(* IEC 61131-3 sources: vespera/src/POU, 15 files *)

(* ---- F_BuildLinks.st ---- *)
(* Связи "кто на кого подаёт" при заданных положениях клапанов.
   Используется для блокировок (с фактическими положениями) и для определения состава
   маршрутов (с положениями из ROUTE_VALVE). Возвращает число связей. *)
FUNCTION F_BuildLinks : INT
VAR_IN_OUT
    aPos   : ARRAY[1..GVL_Const.N_VALVE] OF INT;
    aLinks : ARRAY[1..GVL_Const.N_LINK] OF ST_Link;
END_VAR
VAR
    n : INT;
END_VAR
VAR CONSTANT
    M : INT := 0;   (* LT_MECH *)
    B : INT := 1;   (* LT_BUNKER *)
    X : INT := 2;   (* LT_INVALID *)
END_VAR

(* ---- приёмное отделение и МУЗ ---- *)
n := n + 1; aLinks[n] := F_Link(GVL_Const.M_GATE1, M, GVL_Const.M_N3, TRUE);
n := n + 1; aLinks[n] := F_Link(GVL_Const.M_N3, B, GVL_Const.B_B4, TRUE);
n := n + 1; aLinks[n] := F_Link(GVL_Const.M_MUZ5_FD, M, GVL_Const.M_MUZ5, TRUE);
n := n + 1; aLinks[n] := F_Link(GVL_Const.M_MUZ5, M, GVL_Const.M_N7, TRUE);
n := n + 1; aLinks[n] := F_Link(GVL_Const.M_MUZ5, M, GVL_Const.M_SH32, FALSE);    (* неиспользуемые отходы 32-31-30 *)
n := n + 1; aLinks[n] := F_Link(GVL_Const.M_MUZ5, M, GVL_Const.M_KC35, FALSE);    (* используемые отходы 35-34 *)
n := n + 1; aLinks[n] := F_Link(GVL_Const.M_MUZ5, M, GVL_Const.M_FAN6, FALSE);
n := n + 1; aLinks[n] := F_Link(GVL_Const.M_FAN6, M, GVL_Const.M_SL6, FALSE);
n := n + 1; aLinks[n] := F_Link(GVL_Const.M_N7, B, GVL_Const.B_B8, TRUE);

(* ---- ТОР-18 ---- *)
n := n + 1; aLinks[n] := F_Link(GVL_Const.M_TOR9_FD, M, GVL_Const.M_TOR9, TRUE);
n := n + 1; aLinks[n] := F_Link(GVL_Const.M_TOR9, M, GVL_Const.M_N11, TRUE);
n := n + 1; aLinks[n] := F_Link(GVL_Const.M_TOR9, M, GVL_Const.M_SH31, FALSE);    (* неиспользуемые 31-30 *)
n := n + 1; aLinks[n] := F_Link(GVL_Const.M_TOR9, M, GVL_Const.M_KC35, FALSE);
n := n + 1; aLinks[n] := F_Link(GVL_Const.M_TOR9, M, GVL_Const.M_FAN10, FALSE);
n := n + 1; aLinks[n] := F_Link(GVL_Const.M_FAN10, M, GVL_Const.M_SL10, FALSE);

(* нория 11 -> 12(1) -> TORBA 13(1) | 12(2) -> БТ | растариватель 15(1) -> нория 16 *)
CASE aPos[GVL_Const.V_V12_1] OF
1:
    n := n + 1; aLinks[n] := F_Link(GVL_Const.M_N11, B, GVL_Const.B_T13_1, TRUE);
2:
    CASE aPos[GVL_Const.V_V12_2] OF
    1:
        n := n + 1; aLinks[n] := F_Link(GVL_Const.M_N11, M, GVL_Const.M_BT14_1, TRUE);
        n := n + 1; aLinks[n] := F_Link(GVL_Const.M_N11, M, GVL_Const.M_BT14_2, TRUE);
    2:
        n := n + 1; aLinks[n] := F_Link(GVL_Const.M_N11, M, GVL_Const.M_N16, TRUE);
    ELSE
        n := n + 1; aLinks[n] := F_Link(GVL_Const.M_N11, X, 0, TRUE);
    END_CASE
ELSE
    n := n + 1; aLinks[n] := F_Link(GVL_Const.M_N11, X, 0, TRUE);
END_CASE

(* ---- блок триерный ---- *)
n := n + 1; aLinks[n] := F_Link(GVL_Const.M_BT14_1, M, GVL_Const.M_N16, TRUE);
n := n + 1; aLinks[n] := F_Link(GVL_Const.M_BT14_2, M, GVL_Const.M_N16, TRUE);
n := n + 1; aLinks[n] := F_Link(GVL_Const.M_BT14_1, M, GVL_Const.M_KC36, FALSE);  (* отходы 36-35-34 *)
n := n + 1; aLinks[n] := F_Link(GVL_Const.M_BT14_2, M, GVL_Const.M_KC36, FALSE);

(* нория 16 -> 12(3) -> бункер 17 (КСП) | нория 20 *)
CASE aPos[GVL_Const.V_V12_3] OF
1:
    n := n + 1; aLinks[n] := F_Link(GVL_Const.M_N16, B, GVL_Const.B_B17, TRUE);
2:
    n := n + 1; aLinks[n] := F_Link(GVL_Const.M_N16, M, GVL_Const.M_N20, TRUE);
ELSE
    n := n + 1; aLinks[n] := F_Link(GVL_Const.M_N16, X, 0, TRUE);
END_CASE

(* ---- КСП-11М ---- *)
n := n + 1; aLinks[n] := F_Link(GVL_Const.M_KSP18_FD, M, GVL_Const.M_KSP18, TRUE);
n := n + 1; aLinks[n] := F_Link(GVL_Const.M_KSP18, M, GVL_Const.M_N20, TRUE);
n := n + 1; aLinks[n] := F_Link(GVL_Const.M_KSP18, M, GVL_Const.M_SH33, FALSE);   (* неиспользуемые 33-31-30 *)
n := n + 1; aLinks[n] := F_Link(GVL_Const.M_KSP18, M, GVL_Const.M_KC35, FALSE);
n := n + 1; aLinks[n] := F_Link(GVL_Const.M_KSP18, M, GVL_Const.M_FAN19, FALSE);
n := n + 1; aLinks[n] := F_Link(GVL_Const.M_FAN19, M, GVL_Const.M_SL19, FALSE);
n := n + 1; aLinks[n] := F_Link(GVL_Const.M_N20, B, GVL_Const.B_B22, TRUE);

(* нория 21 -> 12(4) -> бункер 22 (СП) | Z-нория 26 *)
CASE aPos[GVL_Const.V_V12_4] OF
1:
    n := n + 1; aLinks[n] := F_Link(GVL_Const.M_N21, B, GVL_Const.B_B22, TRUE);
2:
    n := n + 1; aLinks[n] := F_Link(GVL_Const.M_N21, M, GVL_Const.M_ZN26, TRUE);
ELSE
    n := n + 1; aLinks[n] := F_Link(GVL_Const.M_N21, X, 0, TRUE);
END_CASE

(* ---- СП-200 ---- *)
n := n + 1; aLinks[n] := F_Link(GVL_Const.M_SP24_DRV, M, GVL_Const.M_ZN26, TRUE);
n := n + 1; aLinks[n] := F_Link(GVL_Const.M_SP24_DRV, M, GVL_Const.M_KC36, FALSE);
n := n + 1; aLinks[n] := F_Link(GVL_Const.M_SP24_DRV, M, GVL_Const.M_SP24_FAN, FALSE);
n := n + 1; aLinks[n] := F_Link(GVL_Const.M_SP24_FAN, M, GVL_Const.M_FAN25, FALSE);
n := n + 1; aLinks[n] := F_Link(GVL_Const.M_FAN25, M, GVL_Const.M_SL25, FALSE);

(* Z-нория 26 -> выгрузка включена: TORBA 13(2) | выключена: бункер фотосепаратора *)
CASE aPos[GVL_Const.V_V49] OF
1:
    n := n + 1; aLinks[n] := F_Link(GVL_Const.M_ZN26, B, GVL_Const.B_T13_2, TRUE);
2:
    n := n + 1; aLinks[n] := F_Link(GVL_Const.M_ZN26, B, GVL_Const.B_B27, TRUE);
ELSE
    n := n + 1; aLinks[n] := F_Link(GVL_Const.M_ZN26, X, 0, TRUE);
END_CASE

(* ---- фотосепаратор (отходы - напрямую в рамку Биг-Бег) ---- *)
n := n + 1; aLinks[n] := F_Link(GVL_Const.M_FS27, M, GVL_Const.M_ZN29, TRUE);
n := n + 1; aLinks[n] := F_Link(GVL_Const.M_FS27, M, GVL_Const.M_FAN28, FALSE);
n := n + 1; aLinks[n] := F_Link(GVL_Const.M_FAN28, M, GVL_Const.M_SL28, FALSE);
n := n + 1; aLinks[n] := F_Link(GVL_Const.M_ZN29, B, GVL_Const.B_T13_2, TRUE);

(* ---- конвейеры отходов ---- *)
n := n + 1; aLinks[n] := F_Link(GVL_Const.M_SH32, M, GVL_Const.M_SH31, FALSE);
n := n + 1; aLinks[n] := F_Link(GVL_Const.M_SH33, M, GVL_Const.M_SH31, FALSE);
n := n + 1; aLinks[n] := F_Link(GVL_Const.M_SH31, M, GVL_Const.M_SH30, FALSE);
n := n + 1; aLinks[n] := F_Link(GVL_Const.M_KC36, M, GVL_Const.M_KC35, FALSE);
n := n + 1; aLinks[n] := F_Link(GVL_Const.M_KC35, M, GVL_Const.M_KC34, FALSE);

F_BuildLinks := n;
END_FUNCTION

(* ---- F_Link.st ---- *)
FUNCTION F_Link : ST_Link
VAR_INPUT
    iFrom    : INT;
    eTo      : INT;
    iTo      : INT;
    xProduct : BOOL;
END_VAR
F_Link.iFrom := iFrom;
F_Link.eTo := eTo;
F_Link.iTo := iTo;
F_Link.xProduct := xProduct;
END_FUNCTION

(* ---- F_Sec.st ---- *)
(* Секунды (UINT) -> TIME *)
FUNCTION F_Sec : TIME
VAR_INPUT
    uSec : UINT;
END_VAR
F_Sec := UDINT_TO_TIME(UINT_TO_UDINT(uSec) * 1000);
END_FUNCTION

(* ---- F_SyncUint.st ---- *)
(* Уставка в RETAIN <-> регистр панели.
   Если панель изменила регистр (он отличается от последнего выданного значения) -
   принять новое значение с ограничением, затем выдать уставку обратно в регистр. *)
FUNCTION F_SyncUint : BOOL
VAR_INPUT
    uMax : UINT;
END_VAR
VAR_IN_OUT
    uHmi    : UINT;
    uPar    : UINT;
    uShadow : UINT;
END_VAR
IF uHmi <> uShadow THEN
    uPar := MIN(uHmi, uMax);
    F_SyncUint := TRUE;
END_IF
uHmi := uPar;
uShadow := uPar;
END_FUNCTION

(* ---- F_SyncWord.st ---- *)
FUNCTION F_SyncWord : BOOL
VAR_IN_OUT
    wHmi    : WORD;
    wPar    : WORD;
    wShadow : WORD;
END_VAR
IF wHmi <> wShadow THEN
    wPar := wHmi;
    F_SyncWord := TRUE;
END_IF
wHmi := wPar;
wShadow := wPar;
END_FUNCTION

(* ---- FB_Bunker.st ---- *)
(* Бункер с датчиком верхнего уровня. Полный бункер ставит на паузу подающий участок
   маршрута; после освобождения и задержки uTRestart участок запускается снова. *)
FUNCTION_BLOCK FB_Bunker
VAR_INPUT
    xHasSF : BOOL;
    stIn   : ST_BunkerIn;
END_VAR
VAR_IN_OUT
    stHmi : ST_BunkerHmi;
    stPar : ST_BunkerPar;
END_VAR
VAR_OUTPUT
    xFull     : BOOL;
    xAlarm    : BOOL;
    xNewAlarm : BOOL;
END_VAR
VAR
    xDvu      : BOOL;
    wAct      : WORD;
    wAlm      : WORD;
    wSts      : WORD;
    uShDvu    : UINT;
    uShRst    : UINT;
    wShByp    : WORD;
    tonFull   : TON;
    tonClear  : TON;
END_VAR

F_SyncUint(uMax := 600, uHmi := stHmi.uTDvu, uPar := stPar.uTDvu, uShadow := uShDvu);
F_SyncUint(uMax := GVL_Const.T_MAX_S, uHmi := stHmi.uTRestart, uPar := stPar.uTRestart, uShadow := uShRst);
F_SyncWord(wHmi := stHmi.wBypass, wPar := stPar.wBypass, wShadow := wShByp);

xDvu := stIn.xDVU AND (stPar.wBypass AND GVL_Const.BY_DVU) = 0;
tonFull(IN := xDvu, PT := F_Sec(stPar.uTDvu));
tonClear(IN := NOT xDvu, PT := F_Sec(stPar.uTRestart));
IF tonFull.Q THEN
    xFull := TRUE;
ELSIF tonClear.Q THEN
    xFull := FALSE;
END_IF

wAct := 0;
IF xHasSF AND NOT stIn.xSF THEN
    wAct := wAct OR GVL_Const.BA_SF;
END_IF
xNewAlarm := (wAct AND NOT wAlm) <> 0;
IF GVL.xReset THEN
    wAlm := wAct;
ELSE
    wAlm := wAlm OR wAct;
END_IF
xAlarm := wAlm <> 0;

wSts := 0;
IF stIn.xDVU THEN wSts := wSts OR GVL_Const.BS_DVU; END_IF
IF xFull THEN wSts := wSts OR GVL_Const.BS_FULL; END_IF
IF stIn.xDNU THEN wSts := wSts OR GVL_Const.BS_DNU; END_IF
IF (stPar.wBypass AND GVL_Const.BY_DVU) <> 0 THEN wSts := wSts OR GVL_Const.BS_BYPASS; END_IF
IF xAlarm THEN wSts := wSts OR GVL_Const.BS_ALARM; END_IF
stHmi.wSts := wSts;
stHmi.wAlm := wAlm;
END_FUNCTION_BLOCK

(* ---- FB_Mech.st ---- *)
(* Механизм линии: двигатель прямого пуска, привод с ПЧ, заслонка с ПЧ или фотосепаратор.

   Режимы:
   - автомат (MODE_AUTO): работает по требованию маршрута. Пуск после задержки uTOn,
     когда все последующие механизмы уже работают (пуск от последнего к первому).
     Останов после задержки uTOff, когда нет требования и остановились все подающие
     механизмы (останов от первого к последнему);
   - ручной с панели (MODE_MAN): кнопки Пуск/Стоп, пуск разрешён только при работе
     последующих механизмов и неполных бункерах на выходе;
   - местный (MODE_LOCAL): ключ поста в "ручн.", кнопки поста;
   - наладка: ручной режим при GVL.xSetup - без блокировок и датчиков безопасности
     (кроме защит двигателя, аварийного стопа и аварии ПЧ).
   Переход между режимами безударный: команда работы сохраняется. *)
FUNCTION_BLOCK FB_Mech
VAR_INPUT
    stCfg       : ST_MechCfg;
    stIn        : ST_MechIn;
    xDemand     : BOOL;    (* требование активного маршрута *)
    xPredRun    : BOOL;    (* работает подающий механизм - удерживать в работе *)
    xSuccOkAuto : BOOL;    (* все последующие механизмы работают *)
    xSuccOkMan  : BOOL;    (* то же + бункеры на выходе не полны *)
    xPaused     : BOOL;    (* участок на паузе по ДВУ (для индикации) *)
END_VAR
VAR_IN_OUT
    stHmi : ST_MechHmi;
    stPar : ST_MechPar;
END_VAR
VAR_OUTPUT
    stOut     : ST_MechOut;
    xRun      : BOOL;      (* механизм в работе (для блокировок соседних) *)
    xCmd      : BOOL;      (* команда работы *)
    xReady    : BOOL;      (* готов к пуску в маршруте *)
    xAuto     : BOOL;
    xAlarm    : BOOL;
    xNewAlarm : BOOL;      (* появилась новая авария (один цикл) *)
END_VAR
VAR
    eMode      : INT;
    xManualReq : BOOL;
    xSetupNow  : BOOL;
    xStartReq  : BOOL;
    xStopReq   : BOOL;
    xMotorOn   : BOOL;     (* выход на двигатель был включен (предыдущий цикл) *)
    xSeqTrip   : BOOL;
    xSeqLatch  : BOOL;
    wAct       : WORD;
    wAlm       : WORD;
    xToDue     : BOOL;
    xOpened    : BOOL;
    xClosed    : BOOL;
    xGoOpen    : BOOL;
    xGoClose   : BOOL;
    xMoveBlock : BOOL;
    wSts       : WORD;
    uShTOn     : UINT;
    uShTOff    : UINT;
    uShTo      : UINT;
    wShByp     : WORD;
    tonStart   : TON;
    tonStop    : TON;
    tonDksRun  : TON;
    tonDksLost : TON;
    rtDks      : R_TRIG;
    tonDsl1    : TON;
    tonDsl2    : TON;
    tonDp      : TON;
    tonFb      : TON;
    tonMove    : TON;
    tpReset    : TP;
    rtCmd      : R_TRIG;
    ftCmd      : F_TRIG;
    tpOn       : TP;
    tpOff      : TP;
    rtLocStart : R_TRIG;
END_VAR

(* ---- уставки панель <-> RETAIN ---- *)
F_SyncUint(uMax := GVL_Const.T_MAX_S, uHmi := stHmi.uTOn, uPar := stPar.uTOn, uShadow := uShTOn);
F_SyncUint(uMax := GVL_Const.T_MAX_S, uHmi := stHmi.uTOff, uPar := stPar.uTOff, uShadow := uShTOff);
F_SyncUint(uMax := 60000, uHmi := stHmi.uToInterval, uPar := stPar.uToInterval, uShadow := uShTo);
F_SyncWord(wHmi := stHmi.wBypass, wPar := stPar.wBypass, wShadow := wShByp);

(* ---- команды панели ---- *)
xStartReq := (stHmi.wCmd AND GVL_Const.C_START) <> 0;
xStopReq := (stHmi.wCmd AND GVL_Const.C_STOP) <> 0;
IF (stHmi.wCmd AND GVL_Const.C_RESET_TO) <> 0 THEN
    stPar.udSecSinceTO := 0;
END_IF
stHmi.wCmd := stHmi.wCmd AND NOT (GVL_Const.C_START OR GVL_Const.C_STOP OR GVL_Const.C_RESET_TO);

(* механизм, занятый маршрутом, в ручной режим с панели не переводится *)
IF xDemand THEN
    stHmi.wCmd := stHmi.wCmd AND NOT GVL_Const.C_MANUAL;
END_IF
xManualReq := (stHmi.wCmd AND GVL_Const.C_MANUAL) <> 0;

IF stCfg.xHasLocal AND stIn.xLocal THEN
    eMode := GVL_Const.MODE_LOCAL;
ELSIF xManualReq THEN
    eMode := GVL_Const.MODE_MAN;
ELSE
    eMode := GVL_Const.MODE_AUTO;
END_IF
xSetupNow := GVL.xSetup AND eMode = GVL_Const.MODE_MAN;
xAuto := eMode = GVL_Const.MODE_AUTO;

(* ---- аварии ---- *)
wAct := 0;
IF stCfg.xHasQF AND NOT stIn.xQF THEN
    wAct := wAct OR GVL_Const.A_QF;
END_IF

tonDksRun(IN := xMotorOn AND stCfg.eDks <> GVL_Const.DKS_NONE, PT := F_Sec(GVL_Retain.stGlobPar.uTDksGrace));
rtDks(CLK := stIn.xDKS);
IF stCfg.eDks = GVL_Const.DKS_PULSE THEN
    (* таймер перезапускается каждым фронтом импульса *)
    tonDksLost(IN := tonDksRun.Q AND NOT rtDks.Q,
               PT := UDINT_TO_TIME(UINT_TO_UDINT(GVL_Retain.stGlobPar.uTDksPulse) * 100));
ELSE
    tonDksLost(IN := tonDksRun.Q AND NOT stIn.xDKS,
               PT := UDINT_TO_TIME(UINT_TO_UDINT(GVL_Retain.stGlobPar.uTDksPulse) * 100));
END_IF
IF tonDksLost.Q AND (stPar.wBypass AND GVL_Const.BY_DKS) = 0 THEN
    wAct := wAct OR GVL_Const.A_DKS;
END_IF

(* сбег ленты контролируется и на стоящей нории: пуск со сбежавшей лентой запрещён *)
tonDsl1(IN := stCfg.xHasDSL AND NOT stIn.xDSL1, PT := T#1S);
IF tonDsl1.Q AND (stPar.wBypass AND GVL_Const.BY_DSL1) = 0 THEN
    wAct := wAct OR GVL_Const.A_DSL1;
END_IF
tonDsl2(IN := stCfg.xHasDSL AND NOT stIn.xDSL2, PT := T#1S);
IF tonDsl2.Q AND (stPar.wBypass AND GVL_Const.BY_DSL2) = 0 THEN
    wAct := wAct OR GVL_Const.A_DSL2;
END_IF
tonDp(IN := stCfg.xHasDP AND NOT stIn.xDP, PT := T#2S);
IF tonDp.Q AND (stPar.wBypass AND GVL_Const.BY_DP) = 0 THEN
    wAct := wAct OR GVL_Const.A_DP;
END_IF

IF stCfg.xHasEStop AND NOT stIn.xEStop THEN
    wAct := wAct OR GVL_Const.A_ESTOP;
END_IF
(* местный "Стоп" при работе от панели/маршрута: механизм уже отключен аппаратно *)
IF stCfg.xHasLocal AND NOT stIn.xLocStop AND eMode <> GVL_Const.MODE_LOCAL AND (xCmd OR xDemand) THEN
    wAct := wAct OR GVL_Const.A_LOCSTOP;
END_IF

CASE stCfg.eKind OF
GVL_Const.K_FC:
    IF stIn.xFcFault THEN
        wAct := wAct OR GVL_Const.A_FC;
    END_IF
    tonFb(IN := xMotorOn AND NOT stIn.xFcReady, PT := F_Sec(GVL_Retain.stGlobPar.uTFcFb));
    IF tonFb.Q THEN
        wAct := wAct OR GVL_Const.A_FCFB;
    END_IF
GVL_Const.K_GATE:
    IF stIn.xFcFault THEN
        wAct := wAct OR GVL_Const.A_FC;
    END_IF
    tonMove(IN := stOut.qOpen OR stOut.qClose, PT := F_Sec(GVL_Retain.stGlobPar.uTGateMove));
    IF tonMove.Q THEN
        wAct := wAct OR GVL_Const.A_MOVE;
    END_IF
    IF stIn.xFb1 AND stIn.xFb2 THEN
        wAct := wAct OR GVL_Const.A_POS;
    END_IF
GVL_Const.K_FS:
    IF stIn.xErr THEN
        wAct := wAct OR GVL_Const.A_FSERR;
    END_IF
    tonFb(IN := xCmd AND NOT stIn.xFb1, PT := F_Sec(GVL_Retain.stGlobPar.uTFsStart));
    IF tonFb.Q THEN
        wAct := wAct OR GVL_Const.A_FSFB;
    END_IF
END_CASE

IF xSetupNow THEN
    wAct := wAct AND GVL_Const.A_HARD;
END_IF

(* фиксация аварий до сброса *)
xNewAlarm := (wAct AND NOT wAlm) <> 0;
IF GVL.xReset THEN
    wAlm := wAct;
    xSeqLatch := FALSE;
ELSE
    wAlm := wAlm OR wAct;
END_IF
xAlarm := wAlm <> 0;

(* ---- готовность к работе в маршруте ---- *)
xReady := NOT xAlarm AND xAuto AND GVL.xGlobalOk
    AND (NOT stCfg.xHasLocal OR stIn.xLocStop)
    AND (NOT stCfg.xHasEStop OR stIn.xEStop)
    AND (stCfg.eKind <> GVL_Const.K_FS
         OR (stIn.xFb2 AND (stIn.xAux OR (stPar.wBypass AND GVL_Const.BY_AUX) <> 0)));

(* ---- команда работы ---- *)
rtLocStart(CLK := stIn.xLocStart);
CASE eMode OF
GVL_Const.MODE_AUTO:
    tonStart(IN := xDemand AND xSuccOkAuto AND xReady AND NOT xCmd, PT := F_Sec(stPar.uTOn));
    IF tonStart.Q THEN
        xCmd := TRUE;
        xSeqLatch := FALSE;
    END_IF
    tonStop(IN := xCmd AND NOT xDemand AND NOT xPredRun, PT := F_Sec(stPar.uTOff));
    IF tonStop.Q THEN
        xCmd := FALSE;
    END_IF
    xSeqTrip := NOT xSuccOkAuto;

GVL_Const.MODE_MAN:
    tonStart(IN := FALSE);
    tonStop(IN := FALSE);
    IF xStartReq AND NOT xAlarm AND GVL.xGlobalOk AND (xSuccOkMan OR xSetupNow) THEN
        xCmd := TRUE;
        xSeqLatch := FALSE;
    END_IF
    IF xStopReq THEN
        xCmd := FALSE;
    END_IF
    xSeqTrip := NOT xSuccOkMan AND NOT xSetupNow;

GVL_Const.MODE_LOCAL:
    tonStart(IN := FALSE);
    tonStop(IN := FALSE);
    IF rtLocStart.Q AND NOT xAlarm AND stIn.xLocStop THEN
        xCmd := TRUE;
    END_IF
    IF NOT stIn.xLocStop THEN
        xCmd := FALSE;
    END_IF
    xSeqTrip := FALSE;
END_CASE

(* заслонка управляется в местном и ручном режимах кнопками открыть/закрыть, см. ниже *)
IF stCfg.eKind = GVL_Const.K_GATE AND eMode <> GVL_Const.MODE_AUTO THEN
    xCmd := FALSE;
    xSeqTrip := FALSE;
END_IF

IF xCmd AND xSeqTrip THEN
    xSeqLatch := TRUE;
END_IF
(* аварийный стоп, пожар, фазы, отключение цепи управления - останов сразу, без задержек *)
IF xAlarm OR NOT GVL.xGlobalOk OR xSeqTrip THEN
    xCmd := FALSE;
END_IF

(* ---- исполнительная часть ---- *)
stOut.qRun := FALSE;
stOut.qPower := FALSE;
stOut.qOpen := FALSE;
stOut.qClose := FALSE;
stOut.qEnable := FALSE;
tpReset(IN := GVL.xReset, PT := T#1S);
stOut.qReset := tpReset.Q;
rtCmd(CLK := xCmd);
ftCmd(CLK := xCmd);
tpOn(IN := rtCmd.Q AND stCfg.eKind = GVL_Const.K_FS, PT := T#1S);
tpOff(IN := ftCmd.Q AND stCfg.eKind = GVL_Const.K_FS, PT := T#1S);
stOut.qOn := tpOn.Q;
stOut.qOff := tpOff.Q;
xOpened := stIn.xFb1 AND NOT stIn.xFb2;
xClosed := stIn.xFb2 AND NOT stIn.xFb1;

CASE stCfg.eKind OF
GVL_Const.K_DOL:
    stOut.qRun := xCmd;
    xRun := xCmd;
    xMotorOn := xCmd;

GVL_Const.K_FC:
    stOut.qPower := GVL.xSysOn AND (NOT stCfg.xHasQF OR stIn.xQF);
    stOut.qRun := xCmd AND stOut.qPower;
    xRun := stOut.qRun;
    xMotorOn := stOut.qRun;

GVL_Const.K_GATE:
    stOut.qPower := GVL.xSysOn AND (NOT stCfg.xHasQF OR stIn.xQF);
    CASE eMode OF
    GVL_Const.MODE_AUTO:
        xGoOpen := xCmd;
        xGoClose := NOT xCmd;
    GVL_Const.MODE_MAN:
        xGoOpen := (stHmi.wCmd AND GVL_Const.C_OPEN) <> 0 AND (xSuccOkMan OR xSetupNow);
        xGoClose := (stHmi.wCmd AND GVL_Const.C_CLOSE) <> 0;
    ELSE
        xGoOpen := stIn.xLocOpen AND stIn.xLocStop;
        xGoClose := stIn.xLocClose AND stIn.xLocStop;
    END_CASE
    (* при общей аварии заслонка только закрывается - прекращение подачи продукта *)
    xGoOpen := xGoOpen AND GVL.xGlobalOk;
    (* ход прекращается при аварии привода или концевиков до сброса *)
    xMoveBlock := (wAlm AND (GVL_Const.A_QF OR GVL_Const.A_FC OR GVL_Const.A_MOVE OR GVL_Const.A_POS)) <> 0
        OR NOT stOut.qPower;
    stOut.qOpen := xGoOpen AND NOT xGoClose AND NOT xOpened AND NOT xMoveBlock;
    stOut.qClose := xGoClose AND NOT xGoOpen AND NOT xClosed AND NOT xMoveBlock;
    (* проём не закрыт - продукт может поступать на норию *)
    xRun := stOut.qOpen OR xOpened OR (NOT xClosed AND NOT xAlarm);
    xMotorOn := stOut.qOpen OR stOut.qClose;

GVL_Const.K_FS:
    stOut.qEnable := xCmd AND stIn.xFb1;
    xRun := xCmd AND stIn.xFb1;
    xMotorOn := xRun;
END_CASE

(* ---- моточасы ---- *)
IF xMotorOn AND GVL.xPulse1s THEN
    stPar.udSecTotal := stPar.udSecTotal + 1;
    stPar.udSecSinceTO := stPar.udSecSinceTO + 1;
END_IF
stHmi.uHoursTotal := UDINT_TO_UINT(MIN(stPar.udSecTotal / 3600, 65535));
stHmi.uMinutes := UDINT_TO_UINT((stPar.udSecTotal / 60) MOD 60);
stHmi.uHoursSinceTO := UDINT_TO_UINT(MIN(stPar.udSecSinceTO / 3600, 65535));
xToDue := stPar.uToInterval > 0 AND stPar.udSecSinceTO / 3600 >= UINT_TO_UDINT(stPar.uToInterval);

(* ---- состояние для панели ---- *)
wSts := 0;
IF xRun THEN wSts := wSts OR GVL_Const.S_RUN; END_IF
IF xCmd THEN wSts := wSts OR GVL_Const.S_CMD; END_IF
IF xReady THEN wSts := wSts OR GVL_Const.S_READY; END_IF
IF xAlarm THEN wSts := wSts OR GVL_Const.S_ALARM; END_IF
IF eMode = GVL_Const.MODE_LOCAL THEN wSts := wSts OR GVL_Const.S_LOCAL; END_IF
IF eMode = GVL_Const.MODE_MAN THEN wSts := wSts OR GVL_Const.S_MANUAL; END_IF
IF xSetupNow THEN wSts := wSts OR GVL_Const.S_SETUP; END_IF
IF tonStart.IN AND NOT xCmd THEN wSts := wSts OR GVL_Const.S_STARTING; END_IF
IF tonStop.IN THEN wSts := wSts OR GVL_Const.S_STOPPING; END_IF
IF xDemand THEN wSts := wSts OR GVL_Const.S_DEMAND; END_IF
IF xPaused THEN wSts := wSts OR GVL_Const.S_PAUSE; END_IF
IF xToDue THEN wSts := wSts OR GVL_Const.S_TO_DUE; END_IF
IF xOpened THEN wSts := wSts OR GVL_Const.S_OPENED; END_IF
IF xClosed THEN wSts := wSts OR GVL_Const.S_CLOSED; END_IF
IF xSeqLatch THEN wSts := wSts OR GVL_Const.S_SEQ_TRIP; END_IF
IF xSuccOkMan THEN wSts := wSts OR GVL_Const.S_SUCC_OK; END_IF
stHmi.wSts := wSts;
stHmi.wAlm := wAlm;

IF xAlarm THEN
    stHmi.iState := 4;
ELSIF eMode = GVL_Const.MODE_LOCAL THEN
    stHmi.iState := 5;
ELSIF tonStop.IN THEN
    stHmi.iState := 3;
ELSIF xRun THEN
    stHmi.iState := 2;
ELSIF tonStart.IN THEN
    stHmi.iState := 1;
ELSE
    stHmi.iState := 0;
END_IF
END_FUNCTION_BLOCK

(* ---- FB_Valve.st ---- *)
(* Переключатель потока ППМ-2 с электроприводом (поз.12(1)..12(4)) и
   механизм промежуточной выгрузки Z-нории поз.26 (пневмораспределитель 49YA1/49YA2).
   Выход держится до срабатывания датчика положения. Положение задаёт маршрут;
   в ручном режиме - кнопки панели, если подающий механизм стоит. *)
FUNCTION_BLOCK FB_Valve
VAR_INPUT
    xHasSF  : BOOL;
    stIn    : ST_ValveIn;
    iTarget : INT;      (* 0 - нет задания маршрута, 1/2 - положение *)
    xFlow   : BOOL;     (* подающий механизм работает *)
END_VAR
VAR_IN_OUT
    stHmi : ST_ValveHmi;
    stPar : ST_ValvePar;
END_VAR
VAR_OUTPUT
    stOut     : ST_ValveOut;
    iPos      : INT;    (* 0 - не определено, 1, 2 *)
    xReady    : BOOL;
    xAlarm    : BOOL;
    xNewAlarm : BOOL;
END_VAR
VAR
    iGoal    : INT;
    xManual  : BOOL;
    xReq1    : BOOL;
    xReq2    : BOOL;
    xMove1   : BOOL;
    xMove2   : BOOL;
    wAct     : WORD;
    wAlm     : WORD;
    wSts     : WORD;
    uShMove  : UINT;
    tonMove  : TON;
    tofQ1    : TOF;
    tofQ2    : TOF;
END_VAR

F_SyncUint(uMax := 600, uHmi := stHmi.uTMove, uPar := stPar.uTMove, uShadow := uShMove);

IF stIn.xS1 AND NOT stIn.xS2 THEN
    iPos := 1;
ELSIF stIn.xS2 AND NOT stIn.xS1 THEN
    iPos := 2;
ELSE
    iPos := 0;
END_IF

(* ---- аварии ---- *)
wAct := 0;
IF xHasSF AND NOT stIn.xSF THEN
    wAct := wAct OR GVL_Const.VA_SF;
END_IF
tonMove(IN := stOut.q1 OR stOut.q2, PT := F_Sec(stPar.uTMove));
IF tonMove.Q THEN
    wAct := wAct OR GVL_Const.VA_TIMEOUT;
END_IF
IF stIn.xS1 AND stIn.xS2 THEN
    wAct := wAct OR GVL_Const.VA_BOTH;
END_IF
xNewAlarm := (wAct AND NOT wAlm) <> 0;
IF GVL.xReset THEN
    wAlm := wAct;
ELSE
    wAlm := wAlm OR wAct;
END_IF
xAlarm := wAlm <> 0;

(* ---- задание положения ---- *)
IF iTarget <> 0 THEN
    stHmi.wCmd := stHmi.wCmd AND NOT GVL_Const.VC_MANUAL;
END_IF
xManual := (stHmi.wCmd AND GVL_Const.VC_MANUAL) <> 0;
xReq1 := (stHmi.wCmd AND GVL_Const.VC_POS1) <> 0;
xReq2 := (stHmi.wCmd AND GVL_Const.VC_POS2) <> 0;
stHmi.wCmd := stHmi.wCmd AND NOT (GVL_Const.VC_POS1 OR GVL_Const.VC_POS2);

IF iTarget <> 0 THEN
    iGoal := iTarget;
ELSIF xManual THEN
    IF NOT xFlow OR GVL.xSetup THEN
        IF xReq1 THEN
            iGoal := 1;
        ELSIF xReq2 THEN
            iGoal := 2;
        END_IF
    END_IF
ELSE
    iGoal := 0;
END_IF

xMove1 := iGoal = 1 AND iPos <> 1 AND NOT xAlarm AND GVL.xGlobalOk;
xMove2 := iGoal = 2 AND iPos <> 2 AND NOT xAlarm AND GVL.xGlobalOk;
(* пауза 0,5 с при реверсе привода *)
stOut.q1 := xMove1 AND NOT tofQ2.Q;
stOut.q2 := xMove2 AND NOT tofQ1.Q AND NOT stOut.q1;
tofQ1(IN := stOut.q1, PT := T#500MS);
tofQ2(IN := stOut.q2, PT := T#500MS);

xReady := NOT xAlarm AND NOT xManual;

wSts := 0;
IF iPos = 1 THEN wSts := wSts OR GVL_Const.VS_POS1; END_IF
IF iPos = 2 THEN wSts := wSts OR GVL_Const.VS_POS2; END_IF
IF stOut.q1 OR stOut.q2 THEN wSts := wSts OR GVL_Const.VS_MOVING; END_IF
IF xAlarm THEN wSts := wSts OR GVL_Const.VS_ALARM; END_IF
IF xManual THEN wSts := wSts OR GVL_Const.VS_MANUAL; END_IF
IF iTarget <> 0 THEN wSts := wSts OR GVL_Const.VS_ROUTE; END_IF
IF xFlow THEN wSts := wSts OR GVL_Const.VS_FLOW; END_IF
stHmi.wSts := wSts;
stHmi.wAlm := wAlm;
END_FUNCTION_BLOCK

(* ---- PLC_PRG.st ---- *)
(* Главная программа. Вызывается из задачи MAST (циклическая, 20 мс). *)
PROGRAM PLC_PRG

PRG_Inputs();
PRG_System();
PRG_Topology();
PRG_Routes();
PRG_Mechs();
PRG_Outputs();
END_PROGRAM

(* ---- PRG_Inputs.st ---- *)
(* Сгенерировано gen/gen_io.py. Физические входы -> логические сигналы.
   Полярность датчиков - константы CFG_* в GVL_Const. *)
PROGRAM PRG_Inputs

GVL.xSysOnIn := GVL_IO.DI_SYS_ON;
GVL.aEStopIn[1] := GVL_IO.DI_ESTOP_1;
GVL.aEStopIn[2] := GVL_IO.DI_ESTOP_2;
GVL.aEStopIn[3] := GVL_IO.DI_ESTOP_3;
GVL.aEStopIn[4] := GVL_IO.DI_ESTOP_4;
GVL.aEStopIn[5] := GVL_IO.DI_ESTOP_5;
GVL.aEStopIn[6] := GVL_IO.DI_ESTOP_6;
GVL.aEStopIn[7] := GVL_IO.DI_ESTOP_7;
GVL.aEStopIn[8] := GVL_IO.DI_ESTOP_8;
GVL.aEStopIn[9] := GVL_IO.DI_ESTOP_9;
GVL.aEStopIn[10] := GVL_IO.DI_ESTOP_10;
GVL.xFireOkIn := GVL_IO.DI_FIRE_OK;
GVL.xPhaseOkIn := GVL_IO.DI_PHASE_OK;
GVL.aMechIn[GVL_Const.M_N3].xDKS := GVL_IO.DI_N3_DKS;
GVL.aMechIn[GVL_Const.M_N3].xDSL1 := (GVL_IO.DI_N3_DSL1 = GVL_Const.CFG_DSL_OK);
GVL.aMechIn[GVL_Const.M_N3].xDSL2 := (GVL_IO.DI_N3_DSL2 = GVL_Const.CFG_DSL_OK);
GVL.aMechIn[GVL_Const.M_N3].xDP := (GVL_IO.DI_N3_DP = GVL_Const.CFG_DP_OK);
GVL.aMechIn[GVL_Const.M_N3].xLocal := (GVL_IO.DI_N3_SA = GVL_Const.CFG_SA_LOCAL);
GVL.aMechIn[GVL_Const.M_N3].xLocStart := GVL_IO.DI_N3_SB_START;
GVL.aMechIn[GVL_Const.M_N3].xLocStop := GVL_IO.DI_N3_SB_STOP;
GVL.aMechIn[GVL_Const.M_N3].xEStop := GVL_IO.DI_N3_SB_ESTOP;
GVL.aMechIn[GVL_Const.M_N3].xQF := GVL_IO.DI_N3_QF;
GVL.aBunkerIn[GVL_Const.B_B4].xDVU := (GVL_IO.DI_B4_DVU = GVL_Const.CFG_DVU_FULL);
GVL.aBunkerIn[GVL_Const.B_B4].xDNU := (GVL_IO.DI_B4_DNU = GVL_Const.CFG_DNU_ON);
GVL.aMechIn[GVL_Const.M_MUZ5].xQF := GVL_IO.DI_MUZ5_QF;
GVL.aMechIn[GVL_Const.M_MUZ5_FD].xQF := GVL_IO.DI_MUZ5FD_SF;
GVL.aMechIn[GVL_Const.M_MUZ5_FD].xFcFault := (GVL_IO.DI_MUZ5FD_FAULT = GVL_Const.CFG_FC_FAULT);
GVL.aMechIn[GVL_Const.M_MUZ5_FD].xFcReady := GVL_IO.DI_MUZ5FD_READY;
GVL.aMechIn[GVL_Const.M_MUZ5_FD].xEStop := GVL_IO.DI_MUZ5FD_ESTOP;
GVL.aMechIn[GVL_Const.M_FAN6].xQF := GVL_IO.DI_FAN6_QF;
GVL.aMechIn[GVL_Const.M_SL6].xDKS := GVL_IO.DI_SL6_DKS;
GVL.aMechIn[GVL_Const.M_SL6].xQF := GVL_IO.DI_SL6_QF;
GVL.aMechIn[GVL_Const.M_N7].xDKS := GVL_IO.DI_N7_DKS;
GVL.aMechIn[GVL_Const.M_N7].xDSL1 := (GVL_IO.DI_N7_DSL1 = GVL_Const.CFG_DSL_OK);
GVL.aMechIn[GVL_Const.M_N7].xDSL2 := (GVL_IO.DI_N7_DSL2 = GVL_Const.CFG_DSL_OK);
GVL.aMechIn[GVL_Const.M_N7].xDP := (GVL_IO.DI_N7_DP = GVL_Const.CFG_DP_OK);
GVL.aMechIn[GVL_Const.M_N7].xLocal := (GVL_IO.DI_N7_SA = GVL_Const.CFG_SA_LOCAL);
GVL.aMechIn[GVL_Const.M_N7].xLocStart := GVL_IO.DI_N7_SB_START;
GVL.aMechIn[GVL_Const.M_N7].xLocStop := GVL_IO.DI_N7_SB_STOP;
GVL.aMechIn[GVL_Const.M_N7].xEStop := GVL_IO.DI_N7_SB_ESTOP;
GVL.aMechIn[GVL_Const.M_N7].xQF := GVL_IO.DI_N7_QF;
GVL.aBunkerIn[GVL_Const.B_B8].xDVU := (GVL_IO.DI_B8_DVU = GVL_Const.CFG_DVU_FULL);
GVL.aBunkerIn[GVL_Const.B_B8].xDNU := (GVL_IO.DI_B8_DNU = GVL_Const.CFG_DNU_ON);
GVL.aMechIn[GVL_Const.M_TOR9].xQF := GVL_IO.DI_TOR9_QF;
GVL.aMechIn[GVL_Const.M_TOR9_FD].xQF := GVL_IO.DI_TOR9FD_SF;
GVL.aMechIn[GVL_Const.M_TOR9_FD].xFcFault := (GVL_IO.DI_TOR9FD_FAULT = GVL_Const.CFG_FC_FAULT);
GVL.aMechIn[GVL_Const.M_TOR9_FD].xFcReady := GVL_IO.DI_TOR9FD_READY;
GVL.aMechIn[GVL_Const.M_TOR9_FD].xEStop := GVL_IO.DI_TOR9FD_ESTOP;
GVL.aMechIn[GVL_Const.M_FAN10].xQF := GVL_IO.DI_FAN10_QF;
GVL.aMechIn[GVL_Const.M_SL10].xDKS := GVL_IO.DI_SL10_DKS;
GVL.aMechIn[GVL_Const.M_SL10].xQF := GVL_IO.DI_SL10_QF;
GVL.aMechIn[GVL_Const.M_N11].xDKS := GVL_IO.DI_N11_DKS;
GVL.aMechIn[GVL_Const.M_N11].xDSL1 := (GVL_IO.DI_N11_DSL1 = GVL_Const.CFG_DSL_OK);
GVL.aMechIn[GVL_Const.M_N11].xDSL2 := (GVL_IO.DI_N11_DSL2 = GVL_Const.CFG_DSL_OK);
GVL.aMechIn[GVL_Const.M_N11].xDP := (GVL_IO.DI_N11_DP = GVL_Const.CFG_DP_OK);
GVL.aMechIn[GVL_Const.M_N11].xLocal := (GVL_IO.DI_N11_SA = GVL_Const.CFG_SA_LOCAL);
GVL.aMechIn[GVL_Const.M_N11].xLocStart := GVL_IO.DI_N11_SB_START;
GVL.aMechIn[GVL_Const.M_N11].xLocStop := GVL_IO.DI_N11_SB_STOP;
GVL.aMechIn[GVL_Const.M_N11].xEStop := GVL_IO.DI_N11_SB_ESTOP;
GVL.aMechIn[GVL_Const.M_N11].xQF := GVL_IO.DI_N11_QF;
GVL.aValveIn[GVL_Const.V_V12_1].xSF := GVL_IO.DI_V121_SF;
GVL.aValveIn[GVL_Const.V_V12_1].xS1 := GVL_IO.DI_V121_POS1;
GVL.aValveIn[GVL_Const.V_V12_1].xS2 := GVL_IO.DI_V121_POS2;
GVL.aValveIn[GVL_Const.V_V12_2].xSF := GVL_IO.DI_V122_SF;
GVL.aValveIn[GVL_Const.V_V12_2].xS1 := GVL_IO.DI_V122_POS1;
GVL.aValveIn[GVL_Const.V_V12_2].xS2 := GVL_IO.DI_V122_POS2;
GVL.aValveIn[GVL_Const.V_V12_3].xSF := GVL_IO.DI_V123_SF;
GVL.aValveIn[GVL_Const.V_V12_3].xS1 := GVL_IO.DI_V123_POS1;
GVL.aValveIn[GVL_Const.V_V12_3].xS2 := GVL_IO.DI_V123_POS2;
GVL.aValveIn[GVL_Const.V_V12_4].xSF := GVL_IO.DI_V124_SF;
GVL.aValveIn[GVL_Const.V_V12_4].xS1 := GVL_IO.DI_V124_POS1;
GVL.aValveIn[GVL_Const.V_V12_4].xS2 := GVL_IO.DI_V124_POS2;
GVL.aBunkerIn[GVL_Const.B_T13_1].xSF := GVL_IO.DI_T131_SF;
GVL.aBunkerIn[GVL_Const.B_T13_2].xSF := GVL_IO.DI_T132_SF;
GVL.aBunkerIn[GVL_Const.B_T13_1].xDVU := (GVL_IO.DI_T131_DVU = GVL_Const.CFG_DVU_FULL);
GVL.aBunkerIn[GVL_Const.B_T13_1].xDNU := (GVL_IO.DI_T131_DNU = GVL_Const.CFG_DNU_ON);
GVL.aBunkerIn[GVL_Const.B_T13_2].xDVU := (GVL_IO.DI_T132_DVU = GVL_Const.CFG_DVU_FULL);
GVL.aBunkerIn[GVL_Const.B_T13_2].xDNU := (GVL_IO.DI_T132_DNU = GVL_Const.CFG_DNU_ON);
GVL.aMechIn[GVL_Const.M_BT14_1].xQF := GVL_IO.DI_BT141_SF;
GVL.aMechIn[GVL_Const.M_BT14_1].xFcFault := (GVL_IO.DI_BT141_FAULT = GVL_Const.CFG_FC_FAULT);
GVL.aMechIn[GVL_Const.M_BT14_1].xFcReady := GVL_IO.DI_BT141_READY;
GVL.aMechIn[GVL_Const.M_BT14_1].xEStop := GVL_IO.DI_BT14_ESTOP;
GVL.aMechIn[GVL_Const.M_BT14_2].xEStop := GVL_IO.DI_BT14_ESTOP;
GVL.aMechIn[GVL_Const.M_BT14_2].xQF := GVL_IO.DI_BT142_SF;
GVL.aMechIn[GVL_Const.M_BT14_2].xFcFault := (GVL_IO.DI_BT142_FAULT = GVL_Const.CFG_FC_FAULT);
GVL.aMechIn[GVL_Const.M_BT14_2].xFcReady := GVL_IO.DI_BT142_READY;
GVL.aMechIn[GVL_Const.M_N16].xDKS := GVL_IO.DI_N16_DKS;
GVL.aMechIn[GVL_Const.M_N16].xDSL1 := (GVL_IO.DI_N16_DSL1 = GVL_Const.CFG_DSL_OK);
GVL.aMechIn[GVL_Const.M_N16].xDSL2 := (GVL_IO.DI_N16_DSL2 = GVL_Const.CFG_DSL_OK);
GVL.aMechIn[GVL_Const.M_N16].xDP := (GVL_IO.DI_N16_DP = GVL_Const.CFG_DP_OK);
GVL.aMechIn[GVL_Const.M_N16].xLocal := (GVL_IO.DI_N16_SA = GVL_Const.CFG_SA_LOCAL);
GVL.aMechIn[GVL_Const.M_N16].xLocStart := GVL_IO.DI_N16_SB_START;
GVL.aMechIn[GVL_Const.M_N16].xLocStop := GVL_IO.DI_N16_SB_STOP;
GVL.aMechIn[GVL_Const.M_N16].xEStop := GVL_IO.DI_N16_SB_ESTOP;
GVL.aMechIn[GVL_Const.M_N16].xQF := GVL_IO.DI_N16_QF;
GVL.aBunkerIn[GVL_Const.B_B17].xDVU := (GVL_IO.DI_B17_DVU = GVL_Const.CFG_DVU_FULL);
GVL.aBunkerIn[GVL_Const.B_B17].xDNU := (GVL_IO.DI_B17_DNU = GVL_Const.CFG_DNU_ON);
GVL.aMechIn[GVL_Const.M_KSP18].xQF := GVL_IO.DI_KSP18_QF;
GVL.aMechIn[GVL_Const.M_KSP18_FD].xQF := GVL_IO.DI_KSP18FD_SF;
GVL.aMechIn[GVL_Const.M_KSP18_FD].xFcFault := (GVL_IO.DI_KSP18FD_FAULT = GVL_Const.CFG_FC_FAULT);
GVL.aMechIn[GVL_Const.M_KSP18_FD].xFcReady := GVL_IO.DI_KSP18FD_READY;
GVL.aMechIn[GVL_Const.M_KSP18_FD].xEStop := GVL_IO.DI_KSP18FD_ESTOP;
GVL.aMechIn[GVL_Const.M_FAN19].xQF := GVL_IO.DI_FAN19_QF;
GVL.aMechIn[GVL_Const.M_SL19].xDKS := GVL_IO.DI_SL19_DKS;
GVL.aMechIn[GVL_Const.M_SL19].xQF := GVL_IO.DI_SL19_QF;
GVL.aMechIn[GVL_Const.M_N20].xDKS := GVL_IO.DI_N20_DKS;
GVL.aMechIn[GVL_Const.M_N20].xDSL1 := (GVL_IO.DI_N20_DSL1 = GVL_Const.CFG_DSL_OK);
GVL.aMechIn[GVL_Const.M_N20].xDSL2 := (GVL_IO.DI_N20_DSL2 = GVL_Const.CFG_DSL_OK);
GVL.aMechIn[GVL_Const.M_N20].xDP := (GVL_IO.DI_N20_DP = GVL_Const.CFG_DP_OK);
GVL.aMechIn[GVL_Const.M_N20].xLocal := (GVL_IO.DI_N20_SA = GVL_Const.CFG_SA_LOCAL);
GVL.aMechIn[GVL_Const.M_N20].xLocStart := GVL_IO.DI_N20_SB_START;
GVL.aMechIn[GVL_Const.M_N20].xLocStop := GVL_IO.DI_N20_SB_STOP;
GVL.aMechIn[GVL_Const.M_N20].xEStop := GVL_IO.DI_N20_SB_ESTOP;
GVL.aMechIn[GVL_Const.M_N20].xQF := GVL_IO.DI_N20_QF;
GVL.aMechIn[GVL_Const.M_N21].xDKS := GVL_IO.DI_N21_DKS;
GVL.aMechIn[GVL_Const.M_N21].xDSL1 := (GVL_IO.DI_N21_DSL1 = GVL_Const.CFG_DSL_OK);
GVL.aMechIn[GVL_Const.M_N21].xDSL2 := (GVL_IO.DI_N21_DSL2 = GVL_Const.CFG_DSL_OK);
GVL.aMechIn[GVL_Const.M_N21].xDP := (GVL_IO.DI_N21_DP = GVL_Const.CFG_DP_OK);
GVL.aMechIn[GVL_Const.M_N21].xLocal := (GVL_IO.DI_N21_SA = GVL_Const.CFG_SA_LOCAL);
GVL.aMechIn[GVL_Const.M_N21].xLocStart := GVL_IO.DI_N21_SB_START;
GVL.aMechIn[GVL_Const.M_N21].xLocStop := GVL_IO.DI_N21_SB_STOP;
GVL.aMechIn[GVL_Const.M_N21].xEStop := GVL_IO.DI_N21_SB_ESTOP;
GVL.aMechIn[GVL_Const.M_N21].xQF := GVL_IO.DI_N21_QF;
GVL.aBunkerIn[GVL_Const.B_B22].xDVU := (GVL_IO.DI_B22_DVU = GVL_Const.CFG_DVU_FULL);
GVL.aBunkerIn[GVL_Const.B_B22].xDNU := (GVL_IO.DI_B22_DNU = GVL_Const.CFG_DNU_ON);
GVL.aMechIn[GVL_Const.M_SP24_FAN].xQF := GVL_IO.DI_SP24FAN_QF;
GVL.aMechIn[GVL_Const.M_SP24_DRV].xQF := GVL_IO.DI_SP24DRV_SF;
GVL.aMechIn[GVL_Const.M_SP24_DRV].xFcFault := (GVL_IO.DI_SP24DRV_FAULT = GVL_Const.CFG_FC_FAULT);
GVL.aMechIn[GVL_Const.M_SP24_DRV].xFcReady := GVL_IO.DI_SP24DRV_READY;
GVL.aMechIn[GVL_Const.M_SP24_DRV].xEStop := GVL_IO.DI_SP24DRV_ESTOP;
GVL.aMechIn[GVL_Const.M_FAN25].xQF := GVL_IO.DI_FAN25_QF;
GVL.aMechIn[GVL_Const.M_SL25].xDKS := GVL_IO.DI_SL25_DKS;
GVL.aMechIn[GVL_Const.M_SL25].xQF := GVL_IO.DI_SL25_QF;
GVL.aMechIn[GVL_Const.M_FAN28].xQF := GVL_IO.DI_FAN28_QF;
GVL.aMechIn[GVL_Const.M_SL28].xDKS := GVL_IO.DI_SL28_DKS;
GVL.aMechIn[GVL_Const.M_SL28].xQF := GVL_IO.DI_SL28_QF;
GVL.aMechIn[GVL_Const.M_SH31].xDKS := GVL_IO.DI_SH31_DKS;
GVL.aMechIn[GVL_Const.M_SH31].xDP := (GVL_IO.DI_SH31_DP = GVL_Const.CFG_DP_SCREW_OK);
GVL.aMechIn[GVL_Const.M_SH31].xLocal := (GVL_IO.DI_SH31_SA = GVL_Const.CFG_SA_LOCAL);
GVL.aMechIn[GVL_Const.M_SH31].xLocStart := GVL_IO.DI_SH31_SB_START;
GVL.aMechIn[GVL_Const.M_SH31].xLocStop := GVL_IO.DI_SH31_SB_STOP;
GVL.aMechIn[GVL_Const.M_SH31].xEStop := GVL_IO.DI_SH31_SB_END;
GVL.aMechIn[GVL_Const.M_SH31].xQF := GVL_IO.DI_SH31_QF;
GVL.aMechIn[GVL_Const.M_SH32].xDKS := GVL_IO.DI_SH32_DKS;
GVL.aMechIn[GVL_Const.M_SH32].xDP := (GVL_IO.DI_SH32_DP = GVL_Const.CFG_DP_SCREW_OK);
GVL.aMechIn[GVL_Const.M_SH32].xLocal := (GVL_IO.DI_SH32_SA = GVL_Const.CFG_SA_LOCAL);
GVL.aMechIn[GVL_Const.M_SH32].xLocStart := GVL_IO.DI_SH32_SB_START;
GVL.aMechIn[GVL_Const.M_SH32].xLocStop := GVL_IO.DI_SH32_SB_STOP;
GVL.aMechIn[GVL_Const.M_SH32].xEStop := GVL_IO.DI_SH32_SB_END;
GVL.aMechIn[GVL_Const.M_SH32].xQF := GVL_IO.DI_SH32_QF;
GVL.aMechIn[GVL_Const.M_SH33].xDKS := GVL_IO.DI_SH33_DKS;
GVL.aMechIn[GVL_Const.M_SH33].xDP := (GVL_IO.DI_SH33_DP = GVL_Const.CFG_DP_SCREW_OK);
GVL.aMechIn[GVL_Const.M_SH33].xLocal := (GVL_IO.DI_SH33_SA = GVL_Const.CFG_SA_LOCAL);
GVL.aMechIn[GVL_Const.M_SH33].xLocStart := GVL_IO.DI_SH33_SB_START;
GVL.aMechIn[GVL_Const.M_SH33].xLocStop := GVL_IO.DI_SH33_SB_STOP;
GVL.aMechIn[GVL_Const.M_SH33].xEStop := GVL_IO.DI_SH33_SB_END;
GVL.aMechIn[GVL_Const.M_SH33].xQF := GVL_IO.DI_SH33_QF;
GVL.aMechIn[GVL_Const.M_KC34].xDKS := GVL_IO.DI_KC34_DKS;
GVL.aMechIn[GVL_Const.M_KC34].xDP := (GVL_IO.DI_KC34_DP = GVL_Const.CFG_DP_CHAIN_OK);
GVL.aMechIn[GVL_Const.M_KC34].xLocal := (GVL_IO.DI_KC34_SA = GVL_Const.CFG_SA_LOCAL);
GVL.aMechIn[GVL_Const.M_KC34].xLocStart := GVL_IO.DI_KC34_SB_START;
GVL.aMechIn[GVL_Const.M_KC34].xLocStop := GVL_IO.DI_KC34_SB_STOP;
GVL.aMechIn[GVL_Const.M_KC34].xEStop := GVL_IO.DI_KC34_SB_END;
GVL.aMechIn[GVL_Const.M_KC34].xQF := GVL_IO.DI_KC34_QF;
GVL.aMechIn[GVL_Const.M_KC35].xDKS := GVL_IO.DI_KC35_DKS;
GVL.aMechIn[GVL_Const.M_KC35].xDP := (GVL_IO.DI_KC35_DP = GVL_Const.CFG_DP_CHAIN_OK);
GVL.aMechIn[GVL_Const.M_KC35].xLocal := (GVL_IO.DI_KC35_SA = GVL_Const.CFG_SA_LOCAL);
GVL.aMechIn[GVL_Const.M_KC35].xLocStart := GVL_IO.DI_KC35_SB_START;
GVL.aMechIn[GVL_Const.M_KC35].xLocStop := GVL_IO.DI_KC35_SB_STOP;
GVL.aMechIn[GVL_Const.M_KC35].xEStop := GVL_IO.DI_KC35_SB_END;
GVL.aMechIn[GVL_Const.M_KC35].xQF := GVL_IO.DI_KC35_QF;
GVL.aMechIn[GVL_Const.M_KC36].xDKS := GVL_IO.DI_KC36_DKS;
GVL.aMechIn[GVL_Const.M_KC36].xDP := (GVL_IO.DI_KC36_DP = GVL_Const.CFG_DP_CHAIN_OK);
GVL.aMechIn[GVL_Const.M_KC36].xLocal := (GVL_IO.DI_KC36_SA = GVL_Const.CFG_SA_LOCAL);
GVL.aMechIn[GVL_Const.M_KC36].xLocStart := GVL_IO.DI_KC36_SB_START;
GVL.aMechIn[GVL_Const.M_KC36].xLocStop := GVL_IO.DI_KC36_SB_STOP;
GVL.aMechIn[GVL_Const.M_KC36].xEStop := GVL_IO.DI_KC36_SB_END;
GVL.aMechIn[GVL_Const.M_KC36].xQF := GVL_IO.DI_KC36_QF;
GVL.aMechIn[GVL_Const.M_SH30].xDKS := GVL_IO.DI_SH30_DKS;
GVL.aMechIn[GVL_Const.M_SH30].xDP := (GVL_IO.DI_SH30_DP = GVL_Const.CFG_DP_SCREW_OK);
GVL.aMechIn[GVL_Const.M_SH30].xLocal := (GVL_IO.DI_SH30_SA = GVL_Const.CFG_SA_LOCAL);
GVL.aMechIn[GVL_Const.M_SH30].xLocStart := GVL_IO.DI_SH30_SB_START;
GVL.aMechIn[GVL_Const.M_SH30].xLocStop := GVL_IO.DI_SH30_SB_STOP;
GVL.aMechIn[GVL_Const.M_SH30].xEStop := GVL_IO.DI_SH30_SB_END;
GVL.aMechIn[GVL_Const.M_SH30].xQF := GVL_IO.DI_SH30_QF;
GVL.aMechIn[GVL_Const.M_ZN26].xDKS := GVL_IO.DI_ZN26_DKS;
GVL.aMechIn[GVL_Const.M_ZN26].xLocal := (GVL_IO.DI_ZN26_SA = GVL_Const.CFG_SA_LOCAL);
GVL.aMechIn[GVL_Const.M_ZN26].xLocStart := GVL_IO.DI_ZN26_SB_START;
GVL.aMechIn[GVL_Const.M_ZN26].xLocStop := GVL_IO.DI_ZN26_SB_STOP;
GVL.aMechIn[GVL_Const.M_ZN26].xEStop := GVL_IO.DI_ZN26_SB_END;
GVL.aMechIn[GVL_Const.M_ZN26].xFcFault := (GVL_IO.DI_ZN26_FAULT = GVL_Const.CFG_FC_FAULT);
GVL.aMechIn[GVL_Const.M_ZN26].xFcReady := GVL_IO.DI_ZN26_READY;
GVL.aMechIn[GVL_Const.M_ZN26].xQF := GVL_IO.DI_ZN26_SF;
GVL.aValveIn[GVL_Const.V_V49].xS1 := GVL_IO.DI_V49_ON;
GVL.aValveIn[GVL_Const.V_V49].xS2 := GVL_IO.DI_V49_OFF;
GVL.aMechIn[GVL_Const.M_ZN29].xDKS := GVL_IO.DI_ZN29_DKS;
GVL.aMechIn[GVL_Const.M_ZN29].xLocal := (GVL_IO.DI_ZN29_SA = GVL_Const.CFG_SA_LOCAL);
GVL.aMechIn[GVL_Const.M_ZN29].xLocStart := GVL_IO.DI_ZN29_SB_START;
GVL.aMechIn[GVL_Const.M_ZN29].xLocStop := GVL_IO.DI_ZN29_SB_STOP;
GVL.aMechIn[GVL_Const.M_ZN29].xEStop := GVL_IO.DI_ZN29_SB_END;
GVL.aMechIn[GVL_Const.M_ZN29].xFcFault := (GVL_IO.DI_ZN29_FAULT = GVL_Const.CFG_FC_FAULT);
GVL.aMechIn[GVL_Const.M_ZN29].xFcReady := GVL_IO.DI_ZN29_READY;
GVL.aMechIn[GVL_Const.M_ZN29].xQF := GVL_IO.DI_ZN29_SF;
GVL.aMechIn[GVL_Const.M_GATE1].xFb1 := GVL_IO.DI_GATE1_OPENED;
GVL.aMechIn[GVL_Const.M_GATE1].xFb2 := GVL_IO.DI_GATE1_CLOSED;
GVL.aMechIn[GVL_Const.M_GATE1].xLocal := (GVL_IO.DI_GATE1_SA = GVL_Const.CFG_SA_LOCAL);
GVL.aMechIn[GVL_Const.M_GATE1].xLocOpen := GVL_IO.DI_GATE1_SB_OPEN;
GVL.aMechIn[GVL_Const.M_GATE1].xLocClose := GVL_IO.DI_GATE1_SB_CLOSE;
GVL.aMechIn[GVL_Const.M_GATE1].xLocStop := GVL_IO.DI_GATE1_SB_STOP;
GVL.aMechIn[GVL_Const.M_GATE1].xFcFault := (GVL_IO.DI_GATE1_FAULT = GVL_Const.CFG_FC_FAULT);
GVL.aMechIn[GVL_Const.M_GATE1].xFcReady := GVL_IO.DI_GATE1_READY;
GVL.aMechIn[GVL_Const.M_GATE1].xQF := GVL_IO.DI_GATE1_SF;
GVL.aBunkerIn[GVL_Const.B_B27].xDVU := (GVL_IO.DI_B27_DVU1 = GVL_Const.CFG_DVU_FULL);
GVL.aBunkerIn[GVL_Const.B_B27].xDNU := (GVL_IO.DI_B27_DVU2 = GVL_Const.CFG_DNU_ON);
GVL.xFsAspPwrIn := GVL_IO.DI_FS27_ASP_SF;
GVL.aMechIn[GVL_Const.M_FS27].xQF := GVL_IO.DI_FS27_SF;
GVL.aMechIn[GVL_Const.M_FS27].xFb1 := GVL_IO.DI_FS27_STATUS;
GVL.aMechIn[GVL_Const.M_FS27].xFb2 := GVL_IO.DI_FS27_REMOTE;
GVL.aMechIn[GVL_Const.M_FS27].xErr := GVL_IO.DI_FS27_ERROR;
GVL.xDryerOkIn := GVL_IO.DI_DRYER_SF;
GVL.xComprOkIn := GVL_IO.DI_COMPR_SF;
GVL.xCompr2OkIn := GVL_IO.DI_COMPR2_SF;
END_PROGRAM

(* ---- PRG_Mechs.st ---- *)
(* Вызов бункеров, клапанов и механизмов *)
PROGRAM PRG_Mechs
VAR
    i       : INT;
    aBunker : ARRAY[1..GVL_Const.N_BUNKER] OF FB_Bunker;
    aValve  : ARRAY[1..GVL_Const.N_VALVE] OF FB_Valve;
    aMech   : ARRAY[1..GVL_Const.N_MECH] OF FB_Mech;
    xAny    : BOOL;
    xNew    : BOOL;
END_VAR

xAny := FALSE;
xNew := FALSE;

FOR i := 1 TO GVL_Const.N_BUNKER DO
    aBunker[i](xHasSF := GVL_Const.BUNKER_HAS_SF[i],
               stIn := GVL.aBunkerIn[i],
               stHmi := GVL_HMI.aHmiBunker[i],
               stPar := GVL_Retain.aBunkerPar[i]);
    GVL.aBunkerFull[i] := aBunker[i].xFull;
    GVL.aBunkerAlarm[i] := aBunker[i].xAlarm;
    xAny := xAny OR aBunker[i].xAlarm;
    xNew := xNew OR aBunker[i].xNewAlarm;
END_FOR

FOR i := 1 TO GVL_Const.N_VALVE DO
    aValve[i](xHasSF := GVL_Const.VALVE_HAS_SF[i],
              stIn := GVL.aValveIn[i],
              iTarget := GVL.aValveTarget[i],
              xFlow := GVL.aRun[GVL_Const.VALVE_FEEDER[i]],
              stHmi := GVL_HMI.aHmiValve[i],
              stPar := GVL_Retain.aValvePar[i]);
    GVL.aValveOut[i] := aValve[i].stOut;
    GVL.aValvePos[i] := aValve[i].iPos;
    GVL.aValveReady[i] := aValve[i].xReady;
    GVL.aValveAlarm[i] := aValve[i].xAlarm;
    xAny := xAny OR aValve[i].xAlarm;
    xNew := xNew OR aValve[i].xNewAlarm;
END_FOR

FOR i := 1 TO GVL_Const.N_MECH DO
    aMech[i](stCfg := GVL_Const.MECH_CFG[i],
             stIn := GVL.aMechIn[i],
             xDemand := GVL.aDemand[i],
             xPredRun := GVL.aPredRun[i],
             xSuccOkAuto := GVL.aSuccAuto[i],
             xSuccOkMan := GVL.aSuccMan[i],
             xPaused := GVL.aBlocked[i],
             stHmi := GVL_HMI.aHmiMech[i],
             stPar := GVL_Retain.aMechPar[i]);
    GVL.aMechOut[i] := aMech[i].stOut;
    GVL.aRun[i] := aMech[i].xRun;
    GVL.aReady[i] := aMech[i].xReady;
    GVL.aAuto[i] := aMech[i].xAuto;
    GVL.aAlarm[i] := aMech[i].xAlarm;
    xAny := xAny OR aMech[i].xAlarm;
    xNew := xNew OR aMech[i].xNewAlarm;
END_FOR

GVL.xAnyAlarm := xAny;
GVL.xAnyNewAlarm := xNew;
END_PROGRAM

(* ---- PRG_Outputs.st ---- *)
(* Сгенерировано gen/gen_io.py. Логические команды -> физические выходы. *)
PROGRAM PRG_Outputs

GVL_IO.DO_SIREN := GVL.qSiren;
GVL_IO.DO_LAMP_ALARM := GVL.qLamp;
GVL_IO.DO_N3_RUN := GVL.aMechOut[GVL_Const.M_N3].qRun;
GVL_IO.DO_MUZ5_RUN := GVL.aMechOut[GVL_Const.M_MUZ5].qRun;
GVL_IO.DO_MUZ5FD_POWER := GVL.aMechOut[GVL_Const.M_MUZ5_FD].qPower;
GVL_IO.DO_MUZ5FD_RESET := GVL.aMechOut[GVL_Const.M_MUZ5_FD].qReset;
GVL_IO.DO_MUZ5FD_RUN := GVL.aMechOut[GVL_Const.M_MUZ5_FD].qRun;
GVL_IO.DO_FAN6_RUN := GVL.aMechOut[GVL_Const.M_FAN6].qRun;
GVL_IO.DO_SL6_RUN := GVL.aMechOut[GVL_Const.M_SL6].qRun;
GVL_IO.DO_N7_RUN := GVL.aMechOut[GVL_Const.M_N7].qRun;
GVL_IO.DO_TOR9_RUN := GVL.aMechOut[GVL_Const.M_TOR9].qRun;
GVL_IO.DO_TOR9FD_POWER := GVL.aMechOut[GVL_Const.M_TOR9_FD].qPower;
GVL_IO.DO_TOR9FD_RESET := GVL.aMechOut[GVL_Const.M_TOR9_FD].qReset;
GVL_IO.DO_TOR9FD_RUN := GVL.aMechOut[GVL_Const.M_TOR9_FD].qRun;
GVL_IO.DO_FAN10_RUN := GVL.aMechOut[GVL_Const.M_FAN10].qRun;
GVL_IO.DO_SL10_RUN := GVL.aMechOut[GVL_Const.M_SL10].qRun;
GVL_IO.DO_N11_RUN := GVL.aMechOut[GVL_Const.M_N11].qRun;
GVL_IO.DO_V121_POS1 := GVL.aValveOut[GVL_Const.V_V12_1].q1;
GVL_IO.DO_V121_POS2 := GVL.aValveOut[GVL_Const.V_V12_1].q2;
GVL_IO.DO_V122_POS1 := GVL.aValveOut[GVL_Const.V_V12_2].q1;
GVL_IO.DO_V122_POS2 := GVL.aValveOut[GVL_Const.V_V12_2].q2;
GVL_IO.DO_V123_POS1 := GVL.aValveOut[GVL_Const.V_V12_3].q1;
GVL_IO.DO_V123_POS2 := GVL.aValveOut[GVL_Const.V_V12_3].q2;
GVL_IO.DO_V124_POS1 := GVL.aValveOut[GVL_Const.V_V12_4].q1;
GVL_IO.DO_V124_POS2 := GVL.aValveOut[GVL_Const.V_V12_4].q2;
GVL_IO.DO_A18_Q9_RES := FALSE;
GVL_IO.DO_BT141_POWER := GVL.aMechOut[GVL_Const.M_BT14_1].qPower;
GVL_IO.DO_BT141_RESET := GVL.aMechOut[GVL_Const.M_BT14_1].qReset;
GVL_IO.DO_BT141_RUN := GVL.aMechOut[GVL_Const.M_BT14_1].qRun;
GVL_IO.DO_BT142_POWER := GVL.aMechOut[GVL_Const.M_BT14_2].qPower;
GVL_IO.DO_BT142_RESET := GVL.aMechOut[GVL_Const.M_BT14_2].qReset;
GVL_IO.DO_BT142_RUN := GVL.aMechOut[GVL_Const.M_BT14_2].qRun;
GVL_IO.DO_N16_RUN := GVL.aMechOut[GVL_Const.M_N16].qRun;
GVL_IO.DO_KSP18_RUN := GVL.aMechOut[GVL_Const.M_KSP18].qRun;
GVL_IO.DO_KSP18FD_POWER := GVL.aMechOut[GVL_Const.M_KSP18_FD].qPower;
GVL_IO.DO_KSP18FD_RESET := GVL.aMechOut[GVL_Const.M_KSP18_FD].qReset;
GVL_IO.DO_KSP18FD_RUN := GVL.aMechOut[GVL_Const.M_KSP18_FD].qRun;
GVL_IO.DO_FAN19_RUN := GVL.aMechOut[GVL_Const.M_FAN19].qRun;
GVL_IO.DO_SL19_RUN := GVL.aMechOut[GVL_Const.M_SL19].qRun;
GVL_IO.DO_N20_RUN := GVL.aMechOut[GVL_Const.M_N20].qRun;
GVL_IO.DO_N21_RUN := GVL.aMechOut[GVL_Const.M_N21].qRun;
GVL_IO.DO_SP24FAN_RUN := GVL.aMechOut[GVL_Const.M_SP24_FAN].qRun;
GVL_IO.DO_SP24DRV_POWER := GVL.aMechOut[GVL_Const.M_SP24_DRV].qPower;
GVL_IO.DO_SP24DRV_RESET := GVL.aMechOut[GVL_Const.M_SP24_DRV].qReset;
GVL_IO.DO_SP24DRV_RUN := GVL.aMechOut[GVL_Const.M_SP24_DRV].qRun;
GVL_IO.DO_FAN25_RUN := GVL.aMechOut[GVL_Const.M_FAN25].qRun;
GVL_IO.DO_SL25_RUN := GVL.aMechOut[GVL_Const.M_SL25].qRun;
GVL_IO.DO_FAN28_RUN := GVL.aMechOut[GVL_Const.M_FAN28].qRun;
GVL_IO.DO_SL28_RUN := GVL.aMechOut[GVL_Const.M_SL28].qRun;
GVL_IO.DO_SH31_RUN := GVL.aMechOut[GVL_Const.M_SH31].qRun;
GVL_IO.DO_SH32_RUN := GVL.aMechOut[GVL_Const.M_SH32].qRun;
GVL_IO.DO_SH33_RUN := GVL.aMechOut[GVL_Const.M_SH33].qRun;
GVL_IO.DO_KC34_RUN := GVL.aMechOut[GVL_Const.M_KC34].qRun;
GVL_IO.DO_KC35_RUN := GVL.aMechOut[GVL_Const.M_KC35].qRun;
GVL_IO.DO_KC36_RUN := GVL.aMechOut[GVL_Const.M_KC36].qRun;
GVL_IO.DO_SH30_RUN := GVL.aMechOut[GVL_Const.M_SH30].qRun;
GVL_IO.DO_ZN26_POWER := GVL.aMechOut[GVL_Const.M_ZN26].qPower;
GVL_IO.DO_ZN26_RUN := GVL.aMechOut[GVL_Const.M_ZN26].qRun;
GVL_IO.DO_ZN26_RESET := GVL.aMechOut[GVL_Const.M_ZN26].qReset;
GVL_IO.DO_V49_ON := GVL.aValveOut[GVL_Const.V_V49].q1;
GVL_IO.DO_V49_OFF := GVL.aValveOut[GVL_Const.V_V49].q2;
GVL_IO.DO_ZN29_POWER := GVL.aMechOut[GVL_Const.M_ZN29].qPower;
GVL_IO.DO_ZN29_RUN := GVL.aMechOut[GVL_Const.M_ZN29].qRun;
GVL_IO.DO_ZN29_RESET := GVL.aMechOut[GVL_Const.M_ZN29].qReset;
GVL_IO.DO_GATE1_POWER := GVL.aMechOut[GVL_Const.M_GATE1].qPower;
GVL_IO.DO_GATE1_OPEN := GVL.aMechOut[GVL_Const.M_GATE1].qOpen;
GVL_IO.DO_GATE1_RESET := GVL.aMechOut[GVL_Const.M_GATE1].qReset;
GVL_IO.DO_GATE1_CLOSE := GVL.aMechOut[GVL_Const.M_GATE1].qClose;
GVL_IO.DO_FS27_ON := GVL.aMechOut[GVL_Const.M_FS27].qOn;
GVL_IO.DO_FS27_OFF := GVL.aMechOut[GVL_Const.M_FS27].qOff;
GVL_IO.DO_FS27_ENABLE := GVL.aMechOut[GVL_Const.M_FS27].qEnable;
GVL_IO.DO_A19_Q23_RES := FALSE;
GVL_IO.DO_A19_Q24_RES := FALSE;
END_PROGRAM

(* ---- PRG_Routes.st ---- *)
(* Маршруты (Приложение 5). Пуск: проверка готовности -> предпусковой сигнал ->
   перевод клапанов -> работа (механизмы запускаются от последнего к первому).
   Стоп: снятие требования (останов от первого к последнему с задержками).
   Авария механизма/клапана/бункера маршрута или общая авария - останов маршрута. *)
PROGRAM PRG_Routes
VAR
    xInit     : BOOL;
    r         : INT;
    p         : INT;
    i         : INT;
    v         : INT;
    b         : INT;
    h         : INT;
    k         : INT;
    nL        : INT;
    aPosT     : ARRAY[1..GVL_Const.N_VALVE] OF INT;
    aL        : ARRAY[1..GVL_Const.N_LINK] OF ST_Link;
    aTonPre   : ARRAY[1..GVL_Const.N_ROUTE] OF TON;
    xToggle   : BOOL;
    xStop     : BOOL;
    xConflict : BOOL;
    xFault    : BOOL;
    xBusy     : BOOL;
    xShared   : BOOL;
    xPaused   : BOOL;
    xAllRun   : BOOL;
    xValvesOk : BOOL;
    iBad      : INT;
    wSts      : WORD;
    aNotReady : ARRAY[1..GVL_Const.N_ROUTE] OF BOOL;
END_VAR

(* ---- состав маршрутов: обход связей от головных механизмов при положениях клапанов маршрута ---- *)
IF NOT xInit THEN
    FOR r := 1 TO GVL_Const.N_ROUTE DO
        FOR v := 1 TO GVL_Const.N_VALVE DO
            aPosT[v] := GVL_Const.ROUTE_VALVE[r, v];
        END_FOR
        nL := F_BuildLinks(aPos := aPosT, aLinks := aL);
        FOR i := 1 TO GVL_Const.N_MECH DO
            GVL.aMember[r, i] := FALSE;
        END_FOR
        FOR b := 1 TO GVL_Const.N_BUNKER DO
            GVL.aMemberB[r, b] := FALSE;
        END_FOR
        GVL.aRouteCfgErr[r] := FALSE;
        FOR h := 1 TO GVL_Const.N_HEAD DO
            IF GVL_Const.ROUTE_HEAD[r, h] > 0 THEN
                GVL.aMember[r, GVL_Const.ROUTE_HEAD[r, h]] := TRUE;
            END_IF
        END_FOR
        FOR p := 1 TO GVL_Const.N_MECH DO
            FOR k := 1 TO nL DO
                IF GVL.aMember[r, aL[k].iFrom] THEN
                    CASE aL[k].eTo OF
                    GVL_Const.LT_MECH:
                        GVL.aMember[r, aL[k].iTo] := TRUE;
                    GVL_Const.LT_BUNKER:
                        GVL.aMemberB[r, aL[k].iTo] := TRUE;
                    ELSE
                        GVL.aRouteCfgErr[r] := TRUE;
                    END_CASE
                END_IF
            END_FOR
        END_FOR
    END_FOR
    xInit := TRUE;
END_IF

FOR r := 1 TO GVL_Const.N_ROUTE DO
    xToggle := (GVL_HMI.aHmiRoute[r].wCmd AND GVL_Const.RC_TOGGLE) <> 0;
    xStop := (GVL_HMI.aHmiRoute[r].wCmd AND GVL_Const.RC_STOP) <> 0 OR GVL.xStopAll;
    GVL_HMI.aHmiRoute[r].wCmd := 0;

    xConflict := FALSE;
    FOR p := 1 TO GVL_Const.N_ROUTE DO
        IF p <> r AND GVL_Const.ROUTE_CONFLICT[r, p] AND GVL.aRouteState[p] <> GVL_Const.RST_IDLE THEN
            xConflict := TRUE;
        END_IF
    END_FOR

    xValvesOk := TRUE;
    FOR v := 1 TO GVL_Const.N_VALVE DO
        IF GVL_Const.ROUTE_VALVE[r, v] <> 0 AND GVL.aValvePos[v] <> GVL_Const.ROUTE_VALVE[r, v] THEN
            xValvesOk := FALSE;
        END_IF
    END_FOR

    (* ---- контроль аварий активного маршрута ---- *)
    IF GVL.aRouteState[r] <> GVL_Const.RST_IDLE AND GVL.aRouteState[r] <> GVL_Const.RST_STOPPING THEN
        xFault := NOT GVL.xGlobalOk;
        FOR i := 1 TO GVL_Const.N_MECH DO
            IF GVL.aMember[r, i] AND (GVL.aAlarm[i] OR NOT GVL.aAuto[i]) THEN
                xFault := TRUE;
            END_IF
        END_FOR
        FOR v := 1 TO GVL_Const.N_VALVE DO
            IF GVL_Const.ROUTE_VALVE[r, v] <> 0 AND GVL.aValveAlarm[v] THEN
                xFault := TRUE;
            END_IF
        END_FOR
        FOR b := 1 TO GVL_Const.N_BUNKER DO
            IF GVL.aMemberB[r, b] AND GVL.aBunkerAlarm[b] THEN
                xFault := TRUE;
            END_IF
        END_FOR
        IF GVL.aRouteState[r] = GVL_Const.RST_RUN AND NOT xValvesOk THEN
            xFault := TRUE;
        END_IF
        IF xFault THEN
            GVL.aRouteFault[r] := TRUE;
            GVL.aRouteState[r] := GVL_Const.RST_STOPPING;
        END_IF
    END_IF

    CASE GVL.aRouteState[r] OF
    GVL_Const.RST_IDLE:
        IF GVL.xReset THEN
            GVL.aRouteFault[r] := FALSE;
            aNotReady[r] := FALSE;
        END_IF
        IF xToggle THEN
            iBad := 0;
            IF NOT GVL.xGlobalOk THEN
                iBad := -1;
            ELSIF xConflict THEN
                iBad := -2;
            ELSIF GVL.aRouteCfgErr[r] THEN
                iBad := -3;
            ELSE
                FOR i := GVL_Const.N_MECH TO 1 BY -1 DO
                    IF GVL.aMember[r, i] AND NOT GVL.aReady[i] THEN
                        iBad := i;
                    END_IF
                END_FOR
                IF iBad = 0 THEN
                    FOR v := GVL_Const.N_VALVE TO 1 BY -1 DO
                        IF GVL_Const.ROUTE_VALVE[r, v] <> 0 AND NOT GVL.aValveReady[v] THEN
                            iBad := 100 + v;
                        END_IF
                    END_FOR
                END_IF
                IF iBad = 0 THEN
                    FOR b := GVL_Const.N_BUNKER TO 1 BY -1 DO
                        IF GVL.aMemberB[r, b] AND GVL.aBunkerAlarm[b] THEN
                            iBad := 200 + b;
                        END_IF
                    END_FOR
                END_IF
            END_IF
            GVL_HMI.aHmiRoute[r].iNotReady := iBad;
            aNotReady[r] := iBad <> 0;
            IF iBad = 0 THEN
                GVL.aRouteFault[r] := FALSE;
                GVL.aRouteState[r] := GVL_Const.RST_PRESTART;
            END_IF
        END_IF

    GVL_Const.RST_PRESTART:
        IF xStop OR xToggle THEN
            GVL.aRouteState[r] := GVL_Const.RST_IDLE;
        ELSIF aTonPre[r].Q THEN
            GVL.aRouteState[r] := GVL_Const.RST_VALVES;
        END_IF

    GVL_Const.RST_VALVES:
        IF xStop OR xToggle THEN
            GVL.aRouteState[r] := GVL_Const.RST_STOPPING;
        ELSIF xValvesOk THEN
            GVL.aRouteState[r] := GVL_Const.RST_RUN;
        END_IF

    GVL_Const.RST_RUN:
        IF xStop OR xToggle THEN
            GVL.aRouteState[r] := GVL_Const.RST_STOPPING;
        END_IF

    GVL_Const.RST_STOPPING:
        (* ждать останова всех механизмов маршрута, кроме занятых другим работающим маршрутом *)
        xBusy := FALSE;
        FOR i := 1 TO GVL_Const.N_MECH DO
            IF GVL.aMember[r, i] AND GVL.aRun[i] THEN
                xShared := FALSE;
                FOR p := 1 TO GVL_Const.N_ROUTE DO
                    IF p <> r AND GVL.aRouteState[p] = GVL_Const.RST_RUN AND GVL.aMember[p, i] THEN
                        xShared := TRUE;
                    END_IF
                END_FOR
                IF NOT xShared THEN
                    xBusy := TRUE;
                END_IF
            END_IF
        END_FOR
        IF NOT xBusy THEN
            GVL.aRouteState[r] := GVL_Const.RST_IDLE;
        END_IF
    END_CASE

    aTonPre[r](IN := GVL.aRouteState[r] = GVL_Const.RST_PRESTART,
               PT := F_Sec(GVL_Retain.stGlobPar.uTPreStart));
END_FOR

(* ---- требования к механизмам и клапанам ---- *)
FOR i := 1 TO GVL_Const.N_MECH DO
    GVL.aDemand[i] := FALSE;
    FOR r := 1 TO GVL_Const.N_ROUTE DO
        IF GVL.aRouteState[r] = GVL_Const.RST_RUN AND GVL.aMember[r, i] THEN
            GVL.aDemand[i] := TRUE;
        END_IF
    END_FOR
    GVL.aDemand[i] := GVL.aDemand[i] AND NOT GVL.aBlocked[i];
END_FOR

GVL.xPreStart := FALSE;
FOR v := 1 TO GVL_Const.N_VALVE DO
    GVL.aValveTarget[v] := 0;
END_FOR
FOR r := 1 TO GVL_Const.N_ROUTE DO
    IF GVL.aRouteState[r] = GVL_Const.RST_PRESTART THEN
        GVL.xPreStart := TRUE;
    END_IF
    IF GVL.aRouteState[r] <> GVL_Const.RST_IDLE THEN
        FOR v := 1 TO GVL_Const.N_VALVE DO
            IF GVL_Const.ROUTE_VALVE[r, v] <> 0 THEN
                GVL.aValveTarget[v] := GVL_Const.ROUTE_VALVE[r, v];
            END_IF
        END_FOR
    END_IF
END_FOR

(* ---- состояние для панели ---- *)
FOR r := 1 TO GVL_Const.N_ROUTE DO
    xConflict := FALSE;
    FOR p := 1 TO GVL_Const.N_ROUTE DO
        IF p <> r AND GVL_Const.ROUTE_CONFLICT[r, p] AND GVL.aRouteState[p] <> GVL_Const.RST_IDLE THEN
            xConflict := TRUE;
        END_IF
    END_FOR
    xPaused := FALSE;
    xAllRun := GVL.aRouteState[r] = GVL_Const.RST_RUN;
    FOR i := 1 TO GVL_Const.N_MECH DO
        IF GVL.aMember[r, i] THEN
            IF GVL.aBlocked[i] THEN
                xPaused := TRUE;
            ELSIF NOT GVL.aRun[i] THEN
                xAllRun := FALSE;
            END_IF
        END_IF
    END_FOR
    wSts := 0;
    IF GVL.aRouteState[r] <> GVL_Const.RST_IDLE THEN wSts := wSts OR GVL_Const.RS_ACTIVE; END_IF
    IF GVL.aRouteState[r] = GVL_Const.RST_PRESTART THEN wSts := wSts OR GVL_Const.RS_PRESTART; END_IF
    IF GVL.aRouteState[r] = GVL_Const.RST_VALVES THEN wSts := wSts OR GVL_Const.RS_VALVES; END_IF
    IF GVL.aRouteState[r] = GVL_Const.RST_RUN THEN wSts := wSts OR GVL_Const.RS_RUN; END_IF
    IF GVL.aRouteState[r] = GVL_Const.RST_STOPPING THEN wSts := wSts OR GVL_Const.RS_STOPPING; END_IF
    IF xPaused AND GVL.aRouteState[r] = GVL_Const.RST_RUN THEN wSts := wSts OR GVL_Const.RS_PAUSED; END_IF
    IF GVL.aRouteFault[r] THEN wSts := wSts OR GVL_Const.RS_FAULT; END_IF
    IF aNotReady[r] THEN wSts := wSts OR GVL_Const.RS_NOTREADY; END_IF
    IF xConflict THEN wSts := wSts OR GVL_Const.RS_CONFLICT; END_IF
    IF xAllRun THEN wSts := wSts OR GVL_Const.RS_ALLRUN; END_IF
    GVL_HMI.aHmiRoute[r].wSts := wSts;
    GVL_HMI.aHmiRoute[r].iState := GVL.aRouteState[r];
END_FOR
END_PROGRAM

(* ---- PRG_System.st ---- *)
(* Общие сигналы: цепь управления, аварийные стопы, пожар, контроль фаз, сброс, наладка,
   сирена и лампа "Авария", секундный импульс, уставки по умолчанию. *)
PROGRAM PRG_System
VAR
    i         : INT;
    wAct      : WORD;
    wAlm      : WORD;
    wWarn     : WORD;
    wSts      : WORD;
    xNewG     : BOOL;
    xSirenLatch : BOOL;
    tonSec    : TON;
    tonBlink  : TON;
    xBlinkReq : BOOL;
    uSh       : ARRAY[1..7] OF UINT;
END_VAR

(* ---- уставки по умолчанию при первом запуске / потере RETAIN ---- *)
IF GVL_Retain.uInitMagic <> GVL_Const.RETAIN_MAGIC THEN
    GVL_Retain.stGlobPar.uTPreStart := 10;
    GVL_Retain.stGlobPar.uTDksGrace := 5;
    GVL_Retain.stGlobPar.uTDksPulse := 30;
    GVL_Retain.stGlobPar.uTFcFb := 5;
    GVL_Retain.stGlobPar.uTFsStart := 60;
    GVL_Retain.stGlobPar.uTGateMove := 90;
    GVL_Retain.stGlobPar.uSirenOn := 1;
    FOR i := 1 TO GVL_Const.N_MECH DO
        GVL_Retain.aMechPar[i].uTOn := GVL_Const.MECH_CFG[i].uDefTOn;
        GVL_Retain.aMechPar[i].uTOff := GVL_Const.MECH_CFG[i].uDefTOff;
        GVL_Retain.aMechPar[i].uToInterval := 0;
        GVL_Retain.aMechPar[i].wBypass := 0;
    END_FOR
    FOR i := 1 TO GVL_Const.N_VALVE DO
        GVL_Retain.aValvePar[i].uTMove := 30;
    END_FOR
    FOR i := 1 TO GVL_Const.N_BUNKER DO
        GVL_Retain.aBunkerPar[i].wBypass := 0;
        GVL_Retain.aBunkerPar[i].uTDvu := 3;
        GVL_Retain.aBunkerPar[i].uTRestart := 30;
    END_FOR
    GVL_Retain.uInitMagic := GVL_Const.RETAIN_MAGIC;
END_IF

F_SyncUint(uMax := 600, uHmi := GVL_HMI.stHmiG.uTPreStart, uPar := GVL_Retain.stGlobPar.uTPreStart, uShadow := uSh[1]);
F_SyncUint(uMax := 600, uHmi := GVL_HMI.stHmiG.uTDksGrace, uPar := GVL_Retain.stGlobPar.uTDksGrace, uShadow := uSh[2]);
F_SyncUint(uMax := 600, uHmi := GVL_HMI.stHmiG.uTDksPulse, uPar := GVL_Retain.stGlobPar.uTDksPulse, uShadow := uSh[3]);
F_SyncUint(uMax := 600, uHmi := GVL_HMI.stHmiG.uTFcFb, uPar := GVL_Retain.stGlobPar.uTFcFb, uShadow := uSh[4]);
F_SyncUint(uMax := 600, uHmi := GVL_HMI.stHmiG.uTFsStart, uPar := GVL_Retain.stGlobPar.uTFsStart, uShadow := uSh[5]);
F_SyncUint(uMax := 600, uHmi := GVL_HMI.stHmiG.uTGateMove, uPar := GVL_Retain.stGlobPar.uTGateMove, uShadow := uSh[6]);
F_SyncUint(uMax := 1, uHmi := GVL_HMI.stHmiG.uSirenOn, uPar := GVL_Retain.stGlobPar.uSirenOn, uShadow := uSh[7]);

(* ---- такты ---- *)
tonSec(IN := NOT tonSec.Q, PT := T#1S);
GVL.xPulse1s := tonSec.Q;
tonBlink(IN := NOT tonBlink.Q, PT := T#500MS);
IF tonBlink.Q THEN
    xBlinkReq := NOT xBlinkReq;
END_IF
GVL.xBlink := xBlinkReq;
IF GVL.xPulse1s THEN
    GVL_HMI.stHmiG.uHeartbeat := GVL_HMI.stHmiG.uHeartbeat + 1;
END_IF

(* ---- команды панели ---- *)
GVL.xReset := (GVL_HMI.stHmiG.wCmd AND GVL_Const.G_RESET) <> 0;
GVL.xStopAll := (GVL_HMI.stHmiG.wCmd AND GVL_Const.G_STOPALL) <> 0;
IF (GVL_HMI.stHmiG.wCmd AND GVL_Const.G_MUTE) <> 0 OR GVL.xReset THEN
    xSirenLatch := FALSE;
END_IF
GVL.xSetup := (GVL_HMI.stHmiG.wCmd AND GVL_Const.G_SETUP) <> 0;
GVL_HMI.stHmiG.wCmd := GVL_HMI.stHmiG.wCmd AND NOT (GVL_Const.G_RESET OR GVL_Const.G_MUTE OR GVL_Const.G_STOPALL);

(* ---- общие аварии ---- *)
GVL.xSysOn := GVL.xSysOnIn;
wAct := 0;
FOR i := 1 TO 10 DO
    IF NOT GVL.aEStopIn[i] THEN
        wAct := wAct OR SHL(WORD#1, i - 1);
    END_IF
END_FOR
IF NOT GVL.xFireOkIn THEN
    wAct := wAct OR GVL_Const.GA_FIRE;
END_IF
IF NOT GVL.xPhaseOkIn THEN
    wAct := wAct OR GVL_Const.GA_PHASE;
END_IF
xNewG := (wAct AND NOT wAlm) <> 0;
IF GVL.xReset THEN
    wAlm := wAct;
ELSE
    wAlm := wAlm OR wAct;
END_IF
GVL.xGlobalOk := GVL.xSysOn AND wAlm = 0;

wWarn := 0;
IF NOT GVL.xComprOkIn THEN wWarn := wWarn OR GVL_Const.GW_COMPR; END_IF
IF NOT GVL.xCompr2OkIn THEN wWarn := wWarn OR GVL_Const.GW_COMPR2; END_IF
IF NOT GVL.xDryerOkIn THEN wWarn := wWarn OR GVL_Const.GW_DRYER; END_IF
IF NOT GVL.xFsAspPwrIn THEN wWarn := wWarn OR GVL_Const.GW_FSASP; END_IF
IF NOT GVL.xSysOn THEN wWarn := wWarn OR GVL_Const.GW_SYSOFF; END_IF
(* сжатый воздух нужен фотосепаратору *)
GVL.aMechIn[GVL_Const.M_FS27].xAux := GVL.xComprOkIn;

(* ---- сирена и лампа (GVL.xAnyAlarm / xAnyNewAlarm - от механизмов, предыдущий цикл) ---- *)
IF (xNewG OR GVL.xAnyNewAlarm) AND GVL_Retain.stGlobPar.uSirenOn <> 0 THEN
    xSirenLatch := TRUE;
END_IF
(* предпусковой сигнал - прерывистый, звучит всегда *)
GVL.qSiren := xSirenLatch OR (GVL.xPreStart AND GVL.xBlink);
GVL.qLamp := (GVL.xAnyAlarm OR wAlm <> 0) AND (GVL.xBlink OR NOT xSirenLatch);

wSts := 0;
IF GVL.xSysOn THEN wSts := wSts OR GVL_Const.GS_SYSON; END_IF
IF GVL.xGlobalOk THEN wSts := wSts OR GVL_Const.GS_OK; END_IF
IF GVL.xAnyAlarm OR wAlm <> 0 THEN wSts := wSts OR GVL_Const.GS_ALARM; END_IF
IF GVL.qSiren THEN wSts := wSts OR GVL_Const.GS_SIREN; END_IF
IF GVL.xSetup THEN wSts := wSts OR GVL_Const.GS_SETUP; END_IF
IF GVL.xPreStart THEN wSts := wSts OR GVL_Const.GS_PRESTART; END_IF
GVL_HMI.stHmiG.wSts := wSts;
GVL_HMI.stHmiG.wAlm := wAlm;
GVL_HMI.stHmiG.wWarn := wWarn;
END_PROGRAM

(* ---- PRG_Topology.st ---- *)
(* Блокировки по фактическим положениям клапанов:
   - aSuccAuto/aSuccMan - все механизмы, на которые подаёт данный, работают;
   - aPredRun - работает механизм, подающий на данный (удержание при останове);
   - aBlocked - полный бункер на выходе участка: пауза от бункера назад до головы участка. *)
PROGRAM PRG_Topology
VAR
    i    : INT;
    k    : INT;
    pass : INT;
    xStop : BOOL;
    xChg : BOOL;
END_VAR

GVL.nLinks := F_BuildLinks(aPos := GVL.aValvePos, aLinks := GVL.aLinks);

FOR i := 1 TO GVL_Const.N_MECH DO
    GVL.aSuccAuto[i] := TRUE;
    GVL.aSuccMan[i] := TRUE;
    GVL.aPredRun[i] := FALSE;
    GVL.aBlocked[i] := FALSE;
END_FOR

FOR k := 1 TO GVL.nLinks DO
    CASE GVL.aLinks[k].eTo OF
    GVL_Const.LT_MECH:
        IF NOT GVL.aRun[GVL.aLinks[k].iTo] THEN
            GVL.aSuccAuto[GVL.aLinks[k].iFrom] := FALSE;
            GVL.aSuccMan[GVL.aLinks[k].iFrom] := FALSE;
        END_IF
        IF GVL.aRun[GVL.aLinks[k].iFrom] THEN
            GVL.aPredRun[GVL.aLinks[k].iTo] := TRUE;
        END_IF
    GVL_Const.LT_BUNKER:
        (* в автомате полный бункер обрабатывается паузой участка (aBlocked) *)
        IF GVL.aBunkerFull[GVL.aLinks[k].iTo] OR GVL.aBunkerAlarm[GVL.aLinks[k].iTo] THEN
            GVL.aSuccMan[GVL.aLinks[k].iFrom] := FALSE;
        END_IF
    ELSE
        GVL.aSuccAuto[GVL.aLinks[k].iFrom] := FALSE;
        GVL.aSuccMan[GVL.aLinks[k].iFrom] := FALSE;
    END_CASE
END_FOR

(* пауза распространяется только по связям продукта и не проходит через бункеры *)
FOR pass := 1 TO GVL_Const.N_MECH DO
    xChg := FALSE;
    FOR k := 1 TO GVL.nLinks DO
        IF GVL.aLinks[k].xProduct AND NOT GVL.aBlocked[GVL.aLinks[k].iFrom] THEN
            (* CASE, а не AND: в ST операнды AND вычисляются оба, индекс iTo зависит от типа *)
            xStop := FALSE;
            CASE GVL.aLinks[k].eTo OF
            GVL_Const.LT_BUNKER: xStop := GVL.aBunkerFull[GVL.aLinks[k].iTo];
            GVL_Const.LT_MECH:   xStop := GVL.aBlocked[GVL.aLinks[k].iTo];
            END_CASE
            IF xStop THEN
                GVL.aBlocked[GVL.aLinks[k].iFrom] := TRUE;
                xChg := TRUE;
            END_IF
        END_IF
    END_FOR
    IF NOT xChg THEN
        EXIT;
    END_IF
END_FOR
END_PROGRAM
